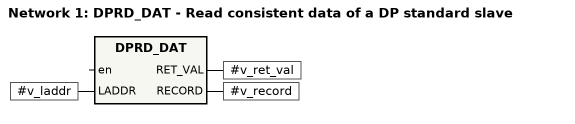
   #v_ret_val := DPRD_DAT(LADDR := #v_laddr, RECORD => #v_record);
END_REGION
END_FUNCTION_BLOCK

FUNCTION_BLOCK "FB_Fbd_ex061"   // FB97, FBD
{ S7_Optimized_Access := 'TRUE' }
   VAR_INPUT
      v_laddr : Hw_Io;
      v_record : Variant;
   END_VAR
   VAR_OUTPUT
      v_ret_val : Int;
   END_VAR
BEGIN

REGION Network 1: DPWR_DAT - Write consistent data of a DP standard slave
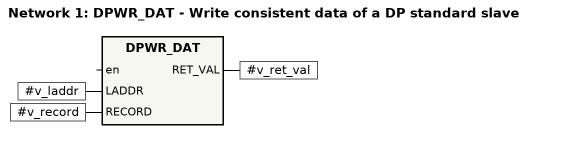
   #v_ret_val := DPWR_DAT(LADDR := #v_laddr, RECORD := #v_record);
END_REGION
END_FUNCTION_BLOCK

FUNCTION_BLOCK "FB_Fbd_ex062"   // FB98, FBD
{ S7_Optimized_Access := 'TRUE' }
   VAR_INPUT
      v_mode : Int;
      v_f_id : Hw_SubModule;
      v_mlen : Int;
      v_code1 : Byte;
      v_code2 : Byte;
   END_VAR
   VAR_OUTPUT
      v_new : Bool;
      v_status : DWord;
      v_slot : Hw_SubModule;
      v_subslot : Hw_SubModule;
      v_index : UInt;
      v_len : UInt;
   END_VAR
   VAR_IN_OUT
      v_record : Array[0..99] of Byte;
   END_VAR
   VAR
      inst : RCVREC;
   END_VAR
BEGIN

REGION Network 1: RCVREC - Receive data record
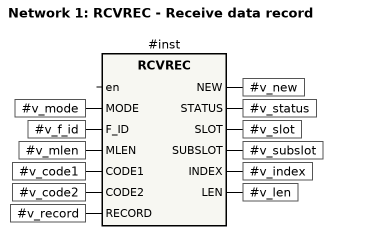
   #inst(MODE := #v_mode,   // RCVREC
         F_ID := #v_f_id,
         MLEN := #v_mlen,
         CODE1 := #v_code1,
         CODE2 := #v_code2,
         RECORD := #v_record,
         NEW => #v_new,
         STATUS => #v_status,
         SLOT => #v_slot,
         SUBSLOT => #v_subslot,
         INDEX => #v_index,
         LEN => #v_len);
END_REGION
END_FUNCTION_BLOCK

FUNCTION_BLOCK "FB_Fbd_ex063"   // FB99, FBD
{ S7_Optimized_Access := 'TRUE' }
   VAR_INPUT
      v_mode : Int;
      v_f_id : Hw_SubModule;
      v_code1 : Byte;
      v_code2 : Byte;
      v_len : UInt;
   END_VAR
   VAR_OUTPUT
      v_new : Bool;
      v_status : DWord;
      v_slot : Hw_SubModule;
      v_subslot : Hw_SubModule;
      v_index : UInt;
      v_rlen : UInt;
   END_VAR
   VAR_IN_OUT
      v_record : Array[0..99] of Byte;
   END_VAR
   VAR
      inst : PRVREC;
   END_VAR
BEGIN

REGION Network 1: PRVREC - Make data record available
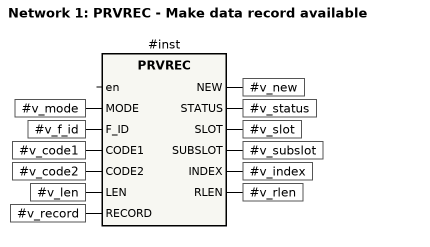
   #inst(MODE := #v_mode,   // PRVREC
         F_ID := #v_f_id,
         CODE1 := #v_code1,
         CODE2 := #v_code2,
         LEN := #v_len,
         RECORD := #v_record,
         NEW => #v_new,
         STATUS => #v_status,
         SLOT => #v_slot,
         SUBSLOT => #v_subslot,
         INDEX => #v_index,
         RLEN => #v_rlen);
END_REGION
END_FUNCTION_BLOCK

FUNCTION_BLOCK "FB_Fbd_ex064"   // FB100, FBD
{ S7_Optimized_Access := 'TRUE' }
   VAR_INPUT
      v_req : Bool;
      v_laddr : Hw_Interface;
      v_group : Byte;
      v_mode : Byte;
   END_VAR
   VAR_OUTPUT
      v_ret_val : Int;
      v_busy : Bool;
   END_VAR
BEGIN

REGION Network 1: DPSYC_FR - Synchronize DP slaves / Freeze inputs
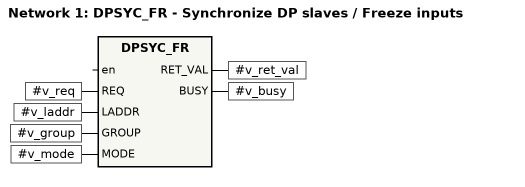
   #v_ret_val := DPSYC_FR(REQ := #v_req, LADDR := #v_laddr, GROUP := #v_group, MODE := #v_mode, BUSY => #v_busy);
END_REGION
END_FUNCTION_BLOCK

FUNCTION_BLOCK "FB_Fbd_ex065"   // FB101, FBD
{ S7_Optimized_Access := 'TRUE' }
   VAR_INPUT
      v_req : Bool;
      v_laddr : Hw_DpSlave;
   END_VAR
   VAR_OUTPUT
      v_ret_val : DInt;
      v_busy : Bool;
   END_VAR
   VAR_IN_OUT
      v_record : Variant;
   END_VAR
BEGIN

REGION Network 1: DPNRM_DG - Read diagnostics data from a DP slave
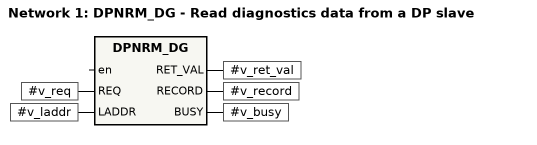
   #v_ret_val := DPNRM_DG(REQ := #v_req, LADDR := #v_laddr, RECORD => #v_record, BUSY => #v_busy);
END_REGION
END_FUNCTION_BLOCK

FUNCTION_BLOCK "FB_Fbd_ex066"   // FB102, FBD
{ S7_Optimized_Access := 'TRUE' }
   VAR_INPUT
      v_req : Bool;
      v_r : Bool;
      v_dp_id : Hw_IoSystem;
   END_VAR
   VAR_OUTPUT
      v_ret_val : Int;
      v_busy : Bool;
      v_dpr : Byte;
      v_dpri : Byte;
   END_VAR
BEGIN

REGION Network 1: DP_TOPOL - Determine topology for DP master system
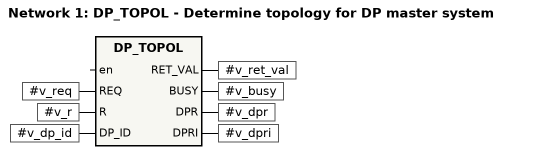
   #v_ret_val := DP_TOPOL(REQ := #v_req,
                          R := #v_r,
                          DP_ID := #v_dp_id,
                          BUSY => #v_busy,
                          DPR => #v_dpr,
                          DPRI => #v_dpri);
END_REGION
END_FUNCTION_BLOCK

FUNCTION_BLOCK "FB_Fbd_ex087"   // FB103, FBD
{ S7_Optimized_Access := 'TRUE' }
   VAR_INPUT
      v_pe_i_dev_new : Bool;
      v_error_code : Byte;
   END_VAR
   VAR_OUTPUT
      v_error : Bool;
      v_status : Word;
   END_VAR
   VAR_IN_OUT
      v_activate : Bool;
      v_valid : Bool;
      v_data_errorrsp : Variant;
   END_VAR
BEGIN

REGION Network 1: PE_Error_RSP - Generate negative answer to command
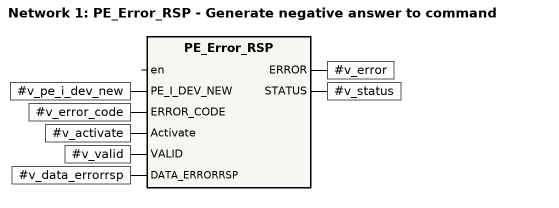
   // no SCL statement known for PE_Error_RSP: written as a call
   PE_Error_RSP(PE_I_DEV_NEW := #v_pe_i_dev_new,
                ERROR_CODE := #v_error_code,
                Activate := #v_activate,
                VALID := #v_valid,
                DATA_ERRORRSP := #v_data_errorrsp,
                ERROR => #v_error,
                STATUS => #v_status);
END_REGION
END_FUNCTION_BLOCK

FUNCTION_BLOCK "FB_Fbd_ex088"   // FB104, FBD
{ S7_Optimized_Access := 'TRUE' }
   VAR_INPUT
      v_pe_i_dev_new : Bool;
      v_cmd : Int;
      v_pe_mode_id : Byte;
   END_VAR
   VAR_OUTPUT
      v_error : Bool;
      v_status : Word;
   END_VAR
   VAR_IN_OUT
      v_activate : Bool;
      v_valid : Bool;
      v_data_errorrsp : Variant;
   END_VAR
BEGIN

REGION Network 1: PE_Start_RSP - Generate answer to command at start of pause
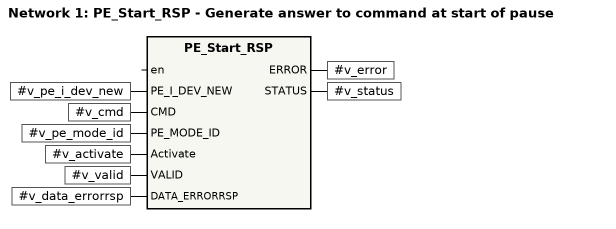
   // no SCL statement known for PE_Start_RSP: written as a call
   PE_Start_RSP(PE_I_DEV_NEW := #v_pe_i_dev_new,
                CMD := #v_cmd,
                PE_MODE_ID := #v_pe_mode_id,
                Activate := #v_activate,
                VALID := #v_valid,
                DATA_ERRORRSP := #v_data_errorrsp,
                ERROR => #v_error,
                STATUS => #v_status);
END_REGION
END_FUNCTION_BLOCK

FUNCTION_BLOCK "FB_Fbd_ex089"   // FB105, FBD
{ S7_Optimized_Access := 'TRUE' }
   VAR_INPUT
      v_pe_i_dev_new : Bool;
      v_cmd : Int;
      v_time_to_operate : DWord;
   END_VAR
   VAR_OUTPUT
      v_error : Bool;
      v_status : Word;
   END_VAR
   VAR_IN_OUT
      v_activate : Bool;
      v_valid : Bool;
      v_data_errorrsp : Variant;
   END_VAR
BEGIN

REGION Network 1: PE_End_RSP - Generate answer to command at end of pause
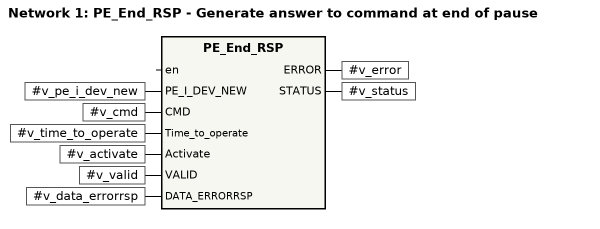
   // no SCL statement known for PE_End_RSP: written as a call
   PE_End_RSP(PE_I_DEV_NEW := #v_pe_i_dev_new,
              CMD := #v_cmd,
              Time_to_operate := #v_time_to_operate,
              Activate := #v_activate,
              VALID := #v_valid,
              DATA_ERRORRSP := #v_data_errorrsp,
              ERROR => #v_error,
              STATUS => #v_status);
END_REGION
END_FUNCTION_BLOCK

FUNCTION_BLOCK "FB_Fbd_ex094"   // FB106, FBD
{ S7_Optimized_Access := 'TRUE' }
   VAR_INPUT
      v_pe_i_dev_new : Bool;
      v_cmd : Int;
      v_cmd_modifier : Int;
      v_count : Byte;
   END_VAR
   VAR_OUTPUT
      v_error : Bool;
      v_status : Word;
   END_VAR
   VAR_IN_OUT
      v_activate : Bool;
      v_valid : Bool;
      v_measurement_list : Variant;
      v_data_errorrsp : Variant;
   END_VAR
BEGIN

REGION Network 1: PE_Measurement_List_RSP - Generate list of supported measured values as answer
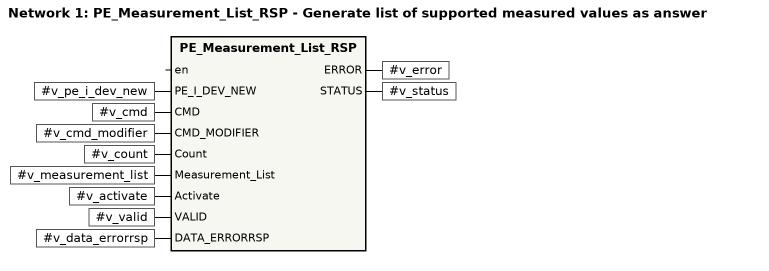
   // no SCL statement known for PE_Measurement_List_RSP: written as a call
   PE_Measurement_List_RSP(PE_I_DEV_NEW := #v_pe_i_dev_new,
                           CMD := #v_cmd,
                           CMD_MODIFIER := #v_cmd_modifier,
                           Count := #v_count,
                           Measurement_List := #v_measurement_list,
                           Activate := #v_activate,
                           VALID := #v_valid,
                           DATA_ERRORRSP := #v_data_errorrsp,
                           ERROR => #v_error,
                           STATUS => #v_status);
END_REGION
END_FUNCTION_BLOCK

FUNCTION_BLOCK "FB_Fbd_ex095"   // FB107, FBD
{ S7_Optimized_Access := 'TRUE' }
   VAR_INPUT
      v_pe_i_dev_new : Bool;
      v_cmd : Int;
      v_cmd_modifier : Int;
      v_count : Byte;
      v_measurement_values : Variant;
   END_VAR
   VAR_OUTPUT
      v_error : Bool;
      v_status : Word;
   END_VAR
   VAR_IN_OUT
      v_activate : Bool;
      v_valid : Bool;
      v_data_errorrsp : Variant;
   END_VAR
BEGIN

REGION Network 1: PE_Measurement_Value_RSP - Generate queried measured values as answer
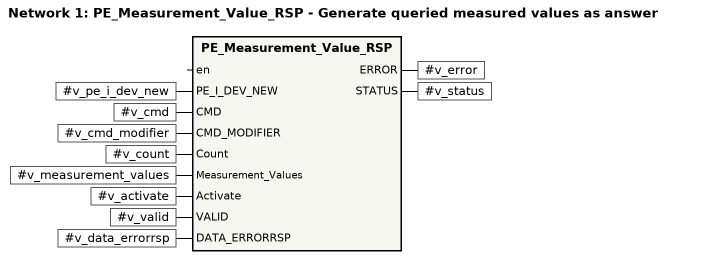
   // no SCL statement known for PE_Measurement_Value_RSP: written as a call
   PE_Measurement_Value_RSP(PE_I_DEV_NEW := #v_pe_i_dev_new,
                           CMD := #v_cmd,
                           CMD_MODIFIER := #v_cmd_modifier,
                           Count := #v_count,
                           Measurement_Values := #v_measurement_values,
                           Activate := #v_activate,
                           VALID := #v_valid,
                           DATA_ERRORRSP := #v_data_errorrsp,
                           ERROR => #v_error,
                           STATUS => #v_status);
END_REGION
END_FUNCTION_BLOCK

FUNCTION_BLOCK "FB_Fbd_ex096"   // FB108, FBD
{ S7_Optimized_Access := 'TRUE' }
   VAR_INPUT
      v_req : Bool;
      v_laddr : Hw_Io;
      v_index : Int;
   END_VAR
   VAR_OUTPUT
      v_valid : Bool;
      v_busy : Bool;
      v_error : Bool;
      v_status : DWord;
      v_len : Int;
   END_VAR
   VAR_IN_OUT
      v_record : Array[0..99] of Byte;
   END_VAR
   VAR
      inst : RD_DPAR;
   END_VAR
BEGIN

REGION Network 1: RD_DPAR - Read module data record
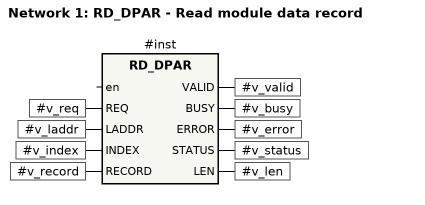
   #inst(REQ := #v_req,   // RD_DPAR
         LADDR := #v_laddr,
         INDEX := #v_index,
         RECORD := #v_record,
         VALID => #v_valid,
         BUSY => #v_busy,
         ERROR => #v_error,
         STATUS => #v_status,
         LEN => #v_len);
END_REGION
END_FUNCTION_BLOCK

FUNCTION_BLOCK "FB_Fbd_ex097"   // FB109, FBD
{ S7_Optimized_Access := 'TRUE' }
   VAR_INPUT
      v_req : Bool;
      v_laddr : Hw_Io;
      v_recnum : Byte;
   END_VAR
   VAR_OUTPUT
      v_ret_val : Int;
      v_busy : Bool;
   END_VAR
   VAR_IN_OUT
      v_record : Variant;
   END_VAR
BEGIN

REGION Network 1: RD_DPARA - Read module data record asynchronously
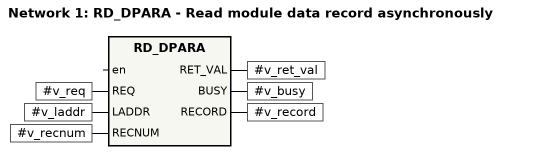
   #v_ret_val := RD_DPARA(REQ := #v_req,
                          LADDR := #v_laddr,
                          RECNUM := #v_recnum,
                          BUSY => #v_busy,
                          RECORD => #v_record);
END_REGION
END_FUNCTION_BLOCK

FUNCTION_BLOCK "FB_Fbd_ex098"   // FB110, FBD
{ S7_Optimized_Access := 'TRUE' }
   VAR_INPUT
      v_ioid : Byte;
      v_laddr : Hw_Io;
      v_recnum : Byte;
   END_VAR
   VAR_OUTPUT
      v_ret_val : Int;
   END_VAR
   VAR_IN_OUT
      v_record : Variant;
   END_VAR
BEGIN

REGION Network 1: RD_DPARM - Read data record from configured system data
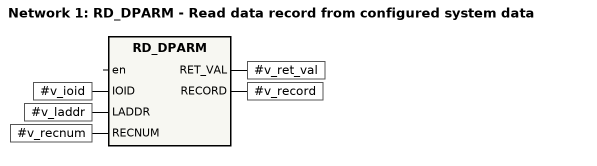
   #v_ret_val := RD_DPARM(IOID := #v_ioid, LADDR := #v_laddr, RECNUM := #v_recnum, RECORD => #v_record);
END_REGION
END_FUNCTION_BLOCK

FUNCTION_BLOCK "FB_Fbd_ex099"   // FB111, FBD
{ S7_Optimized_Access := 'TRUE' }
   VAR_INPUT
      v_req : Bool;
      v_laddr : Hw_Io;
      v_recnum : Byte;
   END_VAR
   VAR_OUTPUT
      v_ret_val : Int;
      v_busy : Bool;
   END_VAR
BEGIN

REGION Network 1: WR_DPARM - Transfer data record
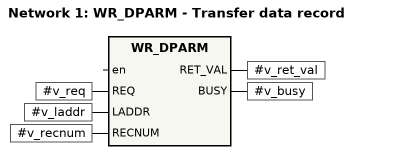
   #v_ret_val := WR_DPARM(REQ := #v_req, LADDR := #v_laddr, RECNUM := #v_recnum, BUSY => #v_busy);
END_REGION
END_FUNCTION_BLOCK

FUNCTION_BLOCK "FB_Fbd_ex100"   // FB112, FBD
{ S7_Optimized_Access := 'TRUE' }
   VAR_INPUT
      v_ob_nr : OB_Att;
      v_event : Event_Att;
      v_add : Bool;
   END_VAR
   VAR_OUTPUT
      v_ret_val : Int;
   END_VAR
BEGIN

REGION Network 1: ATTACH - Attach an OB to an interrupt event
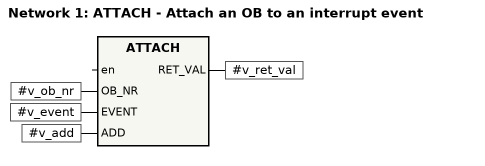
   #v_ret_val := ATTACH(OB_NR := #v_ob_nr, EVENT := #v_event, ADD := #v_add);
END_REGION
END_FUNCTION_BLOCK

FUNCTION_BLOCK "FB_Fbd_ex101"   // FB113, FBD
{ S7_Optimized_Access := 'TRUE' }
   VAR_INPUT
      v_ob_nr : OB_Att;
      v_event : Event_Att;
   END_VAR
   VAR_OUTPUT
      v_ret_val : Int;
   END_VAR
BEGIN

REGION Network 1: DETACH - Detach an OB from an interrupt event
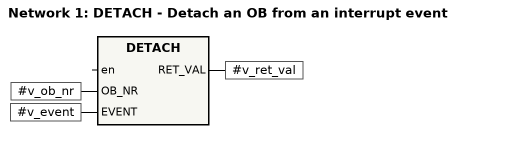
   #v_ret_val := DETACH(OB_NR := #v_ob_nr, EVENT := #v_event);
END_REGION
END_FUNCTION_BLOCK

FUNCTION_BLOCK "FB_Fbd_ex102"   // FB114, FBD
{ S7_Optimized_Access := 'TRUE' }
   VAR_INPUT
      v_ob_nr : OB_Cyclic;
      v_cycle : UDInt;
      v_phase : UDInt;
   END_VAR
   VAR_OUTPUT
      v_ret_val : Int;
   END_VAR
BEGIN

REGION Network 1: SET_CINT - Set cyclic interrupt parameters
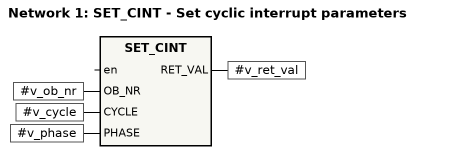
   #v_ret_val := SET_CINT(OB_NR := #v_ob_nr, CYCLE := #v_cycle, PHASE := #v_phase);
END_REGION
END_FUNCTION_BLOCK

FUNCTION_BLOCK "FB_Fbd_ex103"   // FB115, FBD
{ S7_Optimized_Access := 'TRUE' }
   VAR_INPUT
      v_ob_nr : Int;
   END_VAR
   VAR_OUTPUT
      v_cycle : UDInt;
      v_phase : UDInt;
      v_status : Word;
      v_ret_val : Int;
   END_VAR
BEGIN

REGION Network 1: QRY_CINT - Query cyclic interrupt parameters
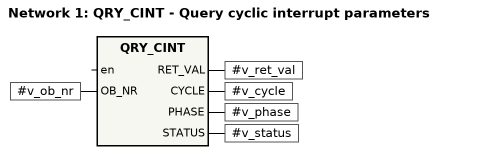
   #v_ret_val := QRY_CINT(OB_NR := #v_ob_nr, CYCLE => #v_cycle, PHASE => #v_phase, STATUS => #v_status);
END_REGION
END_FUNCTION_BLOCK

FUNCTION_BLOCK "FB_Fbd_ex104"   // FB116, FBD
{ S7_Optimized_Access := 'TRUE' }
   VAR_INPUT
      v_ob_nr : OB_Tod;
      v_sdt : Date_And_Time;
      v_period : Word;
   END_VAR
   VAR_OUTPUT
      v_ret_val : Int;
   END_VAR
BEGIN

REGION Network 1: SET_TINT - Set time-of-day interrupt
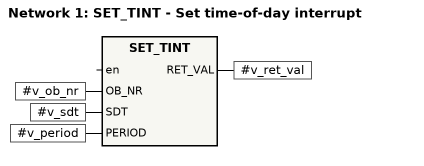
   #v_ret_val := SET_TINT(OB_NR := #v_ob_nr, SDT := #v_sdt, PERIOD := #v_period);
END_REGION
END_FUNCTION_BLOCK

FUNCTION_BLOCK "FB_Fbd_ex105"   // FB117, FBD
{ S7_Optimized_Access := 'TRUE' }
   VAR_INPUT
      v_ob_nr : OB_Tod;
      v_sdt : DTL;
      v_local : Bool;
      v_period : Word;
      v_activate : Bool;
   END_VAR
   VAR_OUTPUT
      v_ret_val : Int;
   END_VAR
BEGIN

REGION Network 1: SET_TINTL - Set time-of-day interrupt
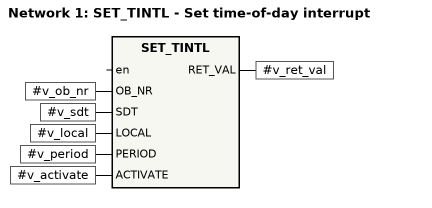
   #v_ret_val := SET_TINTL(OB_NR := #v_ob_nr,
                           SDT := #v_sdt,
                           LOCAL := #v_local,
                           PERIOD := #v_period,
                           ACTIVATE := #v_activate);
END_REGION
END_FUNCTION_BLOCK

FUNCTION_BLOCK "FB_Fbd_ex106"   // FB118, FBD
{ S7_Optimized_Access := 'TRUE' }
   VAR_INPUT
      v_ob_nr : OB_Tod;
   END_VAR
   VAR_OUTPUT
      v_ret_val : Int;
   END_VAR
BEGIN

REGION Network 1: CAN_TINT - Cancel time-of-day interrupt
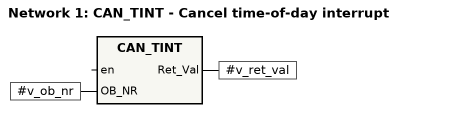
   #v_ret_val := CAN_TINT(OB_NR := #v_ob_nr);
END_REGION
END_FUNCTION_BLOCK

FUNCTION_BLOCK "FB_Fbd_ex107"   // FB119, FBD
{ S7_Optimized_Access := 'TRUE' }
   VAR_INPUT
      v_ob_nr : OB_Tod;
   END_VAR
   VAR_OUTPUT
      v_ret_val : Int;
   END_VAR
BEGIN

REGION Network 1: ACT_TINT - Enable time-of-day interrupt
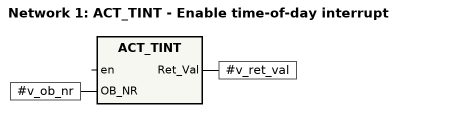
   #v_ret_val := ACT_TINT(OB_NR := #v_ob_nr);
END_REGION
END_FUNCTION_BLOCK

FUNCTION_BLOCK "FB_Fbd_ex108"   // FB120, FBD
{ S7_Optimized_Access := 'TRUE' }
   VAR_INPUT
      v_ob_nr : OB_Tod;
   END_VAR
   VAR_OUTPUT
      v_ret_val : Int;
      v_status : Word;
   END_VAR
BEGIN

REGION Network 1: QRY_TINT - Query status of time-of-day interrupt
